(* IEC 61131-3 sources: plcassist-cli/packages/volt-lsp-iec/test-corpus/bakon-nano/Device/Plc Logic/Application/Library Manager/CAA Storage Imp, 116 files *)

(* ---- _3SSTORAGEVERSIONCONSTANTS.gvl ---- *)
VAR_GLOBAL
	_3SSTORAGE_VERSION_LARGEROREQUAL_3_5_5_0_ : INT := 0;
	_3SSTORAGE_VERSION_LARGEROREQUAL_3_5_11_10_ : INT := 0;
END_VAR

(* ---- GLOBALVARIABLES.gvl ---- *)
VAR_GLOBAL
	FACTORY : StorageFactory;
END_VAR

(* ---- _COLUMNGETBLOB.fun ---- *)
FUNCTION _COLUMNGETBLOB : STO.ERROR
VAR_INPUT
	HROW : ROW;
	IDCOLUMN : CAA.IDENT;
END_VAR
VAR_OUTPUT
	XNULL : BOOL;
END_VAR
VAR_IN_OUT
	BLOBVALUE : STO.STO_BLOB;
END_VAR
END_FUNCTION

(* ---- _COLUMNGETINT16.fun ---- *)
FUNCTION _COLUMNGETINT16 : STO.ERROR
VAR_INPUT
	HROW : ROW;
	IDCOLUMN : CAA.IDENT;
END_VAR
VAR_OUTPUT
	IVALUE : INT;
	XNULL : BOOL;
END_VAR
END_FUNCTION

(* ---- _COLUMNGETINT32.fun ---- *)
FUNCTION _COLUMNGETINT32 : STO.ERROR
VAR_INPUT
	HROW : ROW;
	IDCOLUMN : CAA.IDENT;
END_VAR
VAR_OUTPUT
	DIVALUE : DINT;
	XNULL : BOOL;
END_VAR
END_FUNCTION

(* ---- _COLUMNGETINT64.fun ---- *)
FUNCTION _COLUMNGETINT64 : STO.ERROR
VAR_INPUT
	HROW : ROW;
	IDCOLUMN : CAA.IDENT;
END_VAR
VAR_OUTPUT
	LIVALUE : LINT;
	XNULL : BOOL;
END_VAR
END_FUNCTION

(* ---- _COLUMNGETINT8.fun ---- *)
FUNCTION _COLUMNGETINT8 : STO.ERROR
VAR_INPUT
	HROW : ROW;
	IDCOLUMN : CAA.IDENT;
END_VAR
VAR_OUTPUT
	SIVALUE : SINT;
	XNULL : BOOL;
END_VAR
END_FUNCTION

(* ---- _COLUMNGETREAL4.fun ---- *)
FUNCTION _COLUMNGETREAL4 : STO.ERROR
VAR_INPUT
	HROW : ROW;
	IDCOLUMN : CAA.IDENT;
END_VAR
VAR_OUTPUT
	RVALUE : REAL;
	XNULL : BOOL;
END_VAR
END_FUNCTION

(* ---- _COLUMNGETREAL8.fun ---- *)
FUNCTION _COLUMNGETREAL8 : STO.ERROR
VAR_INPUT
	HROW : ROW;
	IDCOLUMN : CAA.IDENT;
END_VAR
VAR_OUTPUT
	LRVALUE : LREAL;
	XNULL : BOOL;
END_VAR
END_FUNCTION

(* ---- _COLUMNGETTEXT.fun ---- *)
FUNCTION _COLUMNGETTEXT : STO.ERROR
VAR_INPUT
	HROW : ROW;
	IDCOLUMN : CAA.IDENT;
END_VAR
VAR_OUTPUT
	XNULL : BOOL;
END_VAR
VAR_IN_OUT
	TXTVALUE : STO.STO_TEXT;
END_VAR
END_FUNCTION

(* ---- _COLUMNGETTYPE.fun ---- *)
FUNCTION _COLUMNGETTYPE : STO.COLUMN_TYPE
VAR_INPUT
	HROW : ROW;
	IDCOLUMN : CAA.IDENT;
END_VAR
VAR_OUTPUT
	EERROR : STO.ERROR;
END_VAR
END_FUNCTION

(* ---- _COLUMNSETBLOB.fun ---- *)
FUNCTION _COLUMNSETBLOB : STO.ERROR
VAR_INPUT
	HROW : ROW;
	IDCOLUMN : CAA.IDENT;
END_VAR
VAR_IN_OUT
	BLOBVALUE : STO.STO_BLOB;
END_VAR
END_FUNCTION

(* ---- _COLUMNSETINT16.fun ---- *)
FUNCTION _COLUMNSETINT16 : STO.ERROR
VAR_INPUT
	HROW : ROW;
	IDCOLUMN : CAA.IDENT;
	IVALUE : INT;
END_VAR
END_FUNCTION

(* ---- _COLUMNSETINT32.fun ---- *)
FUNCTION _COLUMNSETINT32 : STO.ERROR
VAR_INPUT
	HROW : ROW;
	IDCOLUMN : CAA.IDENT;
	DIVALUE : DINT;
END_VAR
END_FUNCTION

(* ---- _COLUMNSETINT64.fun ---- *)
FUNCTION _COLUMNSETINT64 : STO.ERROR
VAR_INPUT
	HROW : ROW;
	IDCOLUMN : CAA.IDENT;
	LIVALUE : LINT;
END_VAR
END_FUNCTION

(* ---- _COLUMNSETINT8.fun ---- *)
FUNCTION _COLUMNSETINT8 : STO.ERROR
VAR_INPUT
	HROW : ROW;
	IDCOLUMN : CAA.IDENT;
	SIVALUE : SINT;
END_VAR
END_FUNCTION

(* ---- _COLUMNSETNULL.fun ---- *)
FUNCTION _COLUMNSETNULL : STO.ERROR
VAR_INPUT
	HROW : ROW;
	IDCOLUMN : CAA.IDENT;
END_VAR
END_FUNCTION

(* ---- _COLUMNSETREAL4.fun ---- *)
FUNCTION _COLUMNSETREAL4 : STO.ERROR
VAR_INPUT
	HROW : ROW;
	IDCOLUMN : CAA.IDENT;
	RVALUE : REAL;
END_VAR
END_FUNCTION

(* ---- _COLUMNSETREAL8.fun ---- *)
FUNCTION _COLUMNSETREAL8 : STO.ERROR
VAR_INPUT
	HROW : ROW;
	IDCOLUMN : CAA.IDENT;
	LRVALUE : LREAL;
END_VAR
END_FUNCTION

(* ---- _COLUMNSETTEXT.fun ---- *)
FUNCTION _COLUMNSETTEXT : STO.ERROR
VAR_INPUT
	HROW : ROW;
	IDCOLUMN : CAA.IDENT;
END_VAR
VAR_IN_OUT
	TXTVALUE : STO.STO_TEXT;
END_VAR
END_FUNCTION

(* ---- _COLUMNUPDATEBLOB.fun ---- *)
FUNCTION _COLUMNUPDATEBLOB : STO.ERROR
VAR_INPUT
	HROW : ROW;
	IDCOLUMN : CAA.IDENT;
END_VAR
VAR_IN_OUT
	BLOBVALUE : STO.STO_BLOB;
	XNULL : BOOL;
END_VAR
END_FUNCTION

(* ---- _COLUMNUPDATEINT16.fun ---- *)
FUNCTION _COLUMNUPDATEINT16 : STO.ERROR
VAR_INPUT
	HROW : ROW;
	IDCOLUMN : CAA.IDENT;
END_VAR
VAR_IN_OUT
	IVALUE : INT;
	XNULL : BOOL;
END_VAR
END_FUNCTION

(* ---- _COLUMNUPDATEINT32.fun ---- *)
FUNCTION _COLUMNUPDATEINT32 : STO.ERROR
VAR_INPUT
	HROW : ROW;
	IDCOLUMN : CAA.IDENT;
END_VAR
VAR_IN_OUT
	DIVALUE : DINT;
	XNULL : BOOL;
END_VAR
END_FUNCTION

(* ---- _COLUMNUPDATEINT64.fun ---- *)
FUNCTION _COLUMNUPDATEINT64 : STO.ERROR
VAR_INPUT
	HROW : ROW;
	IDCOLUMN : CAA.IDENT;
END_VAR
VAR_IN_OUT
	LIVALUE : LINT;
	XNULL : BOOL;
END_VAR
END_FUNCTION

(* ---- _COLUMNUPDATEINT8.fun ---- *)
FUNCTION _COLUMNUPDATEINT8 : STO.ERROR
VAR_INPUT
	HROW : ROW;
	IDCOLUMN : CAA.IDENT;
END_VAR
VAR_IN_OUT
	SIVALUE : SINT;
	XNULL : BOOL;
END_VAR
END_FUNCTION

(* ---- _COLUMNUPDATEREAL4.fun ---- *)
FUNCTION _COLUMNUPDATEREAL4 : STO.ERROR
VAR_INPUT
	HROW : ROW;
	IDCOLUMN : CAA.IDENT;
END_VAR
VAR_IN_OUT
	RVALUE : REAL;
	XNULL : BOOL;
END_VAR
END_FUNCTION

(* ---- _COLUMNUPDATEREAL8.fun ---- *)
FUNCTION _COLUMNUPDATEREAL8 : STO.ERROR
VAR_INPUT
	HROW : ROW;
	IDCOLUMN : CAA.IDENT;
END_VAR
VAR_IN_OUT
	LRVALUE : LREAL;
	XNULL : BOOL;
END_VAR
END_FUNCTION

(* ---- _COLUMNUPDATETEXT.fun ---- *)
FUNCTION _COLUMNUPDATETEXT : STO.ERROR
VAR_INPUT
	HROW : ROW;
	IDCOLUMN : CAA.IDENT;
END_VAR
VAR_IN_OUT
	TXTVALUE : STO.STO_TEXT;
	XNULL : BOOL;
END_VAR
END_FUNCTION

(* ---- _CURSORCLOSE.fun ---- *)
FUNCTION _CURSORCLOSE : STO.ERROR
VAR_INPUT
	HCURSOR : CURSOR;
END_VAR
END_FUNCTION

(* ---- _CURSORGETCURRENTROW.fun ---- *)
FUNCTION _CURSORGETCURRENTROW : ROW
VAR_INPUT
	HCURSOR : CURSOR;
END_VAR
VAR_OUTPUT
	EERROR : STO.ERROR;
END_VAR
END_FUNCTION

(* ---- _CURSORGETINDEXID.fun ---- *)
FUNCTION _CURSORGETINDEXID : CAA.IDENT
VAR_INPUT
	HCURSOR : CURSOR;
END_VAR
VAR_OUTPUT
	EERROR : STO.ERROR;
END_VAR
END_FUNCTION

(* ---- _CURSORGETSTORAGE.fun ---- *)
FUNCTION _CURSORGETSTORAGE : STORAGE_TYPE
VAR_INPUT
	HCURSOR : CURSOR;
END_VAR
VAR_OUTPUT
	EERROR : STO.ERROR;
END_VAR
END_FUNCTION

(* ---- _CURSORGETTABLE.fun ---- *)
FUNCTION _CURSORGETTABLE : TABLE
VAR_INPUT
	HCURSOR : CURSOR;
END_VAR
VAR_OUTPUT
	EERROR : STO.ERROR;
END_VAR
END_FUNCTION

(* ---- _CURSORISREADONLY.fun ---- *)
FUNCTION _CURSORISREADONLY : BOOL
VAR_INPUT
	HCURSOR : CURSOR;
END_VAR
VAR_OUTPUT
	EERROR : STO.ERROR;
END_VAR
END_FUNCTION

(* ---- _CURSORMOVE.fun ---- *)
FUNCTION _CURSORMOVE : STO.ERROR
VAR_INPUT
	HCURSOR : CURSOR;
	EDIRECTION : STO.DIRECTION;
END_VAR
END_FUNCTION

(* ---- _CURSOROPEN.fun ---- *)
FUNCTION _CURSOROPEN : CURSOR
VAR_INPUT
	HTABLE : TABLE;
	IDINDEX : CAA.IDENT;
	XREADONLY : BOOL;
END_VAR
VAR_OUTPUT
	EERROR : STO.ERROR;
END_VAR
END_FUNCTION

(* ---- _CURSORSEARCHINT16.fun ---- *)
FUNCTION _CURSORSEARCHINT16 : STO.ERROR
VAR_INPUT
	HCURSOR : CURSOR;
	IVALUE : INT;
END_VAR
END_FUNCTION

(* ---- _CURSORSEARCHINT32.fun ---- *)
FUNCTION _CURSORSEARCHINT32 : STO.ERROR
VAR_INPUT
	HCURSOR : CURSOR;
	DIVALUE : DINT;
END_VAR
END_FUNCTION

(* ---- _CURSORSEARCHINT64.fun ---- *)
FUNCTION _CURSORSEARCHINT64 : STO.ERROR
VAR_INPUT
	HCURSOR : CURSOR;
	LIVALUE : LINT;
END_VAR
END_FUNCTION

(* ---- _CURSORSEARCHINT8.fun ---- *)
FUNCTION _CURSORSEARCHINT8 : STO.ERROR
VAR_INPUT
	HCURSOR : CURSOR;
	SIVALUE : SINT;
END_VAR
END_FUNCTION

(* ---- _CURSORSEARCHNULL.fun ---- *)
FUNCTION _CURSORSEARCHNULL : STO.ERROR
VAR_INPUT
	HCURSOR : CURSOR;
END_VAR
END_FUNCTION

(* ---- _CURSORSEARCHREAL4.fun ---- *)
FUNCTION _CURSORSEARCHREAL4 : STO.ERROR
VAR_INPUT
	HCURSOR : CURSOR;
	RVALUE : REAL;
END_VAR
END_FUNCTION

(* ---- _CURSORSEARCHREAL8.fun ---- *)
FUNCTION _CURSORSEARCHREAL8 : STO.ERROR
VAR_INPUT
	HCURSOR : CURSOR;
	LRVALUE : LREAL;
END_VAR
END_FUNCTION

(* ---- _CURSORSEARCHROWID.fun ---- *)
FUNCTION _CURSORSEARCHROWID : STO.ERROR
VAR_INPUT
	HCURSOR : CURSOR;
	IDROW : CAA.IDENT;
END_VAR
END_FUNCTION

(* ---- _CURSORSEARCHROWID2.fun ---- *)
FUNCTION _CURSORSEARCHROWID2 : STO.ERROR
VAR_INPUT
	HCURSOR : CURSOR;
	IDROW : LINT;
END_VAR
END_FUNCTION

(* ---- _CURSORSEARCHTEXT.fun ---- *)
FUNCTION _CURSORSEARCHTEXT : STO.ERROR
VAR_INPUT
	HCURSOR : CURSOR;
END_VAR
VAR_IN_OUT
	TXTVALUE : STO.STO_TEXT;
END_VAR
END_FUNCTION

(* ---- _ROWCLEAR.fun ---- *)
FUNCTION _ROWCLEAR : STO.ERROR
VAR_INPUT
	HROW : ROW;
END_VAR
END_FUNCTION

(* ---- _ROWCREATE.fun ---- *)
FUNCTION _ROWCREATE : ROW
VAR_INPUT
	HTABLE : TABLE;
END_VAR
VAR_OUTPUT
	EERROR : STO.ERROR;
END_VAR
END_FUNCTION

(* ---- _ROWDELETE.fun ---- *)
FUNCTION _ROWDELETE : STO.ERROR
VAR_INPUT
	HTABLE : TABLE;
	IDROW : CAA.IDENT;
END_VAR
END_FUNCTION

(* ---- _ROWDELETE2.fun ---- *)
FUNCTION _ROWDELETE2 : STO.ERROR
VAR_INPUT
	HTABLE : TABLE;
	IDROW : LINT;
END_VAR
END_FUNCTION

(* ---- _ROWDUPLICATE.fun ---- *)
FUNCTION _ROWDUPLICATE : ROW
VAR_INPUT
	HTABLE : TABLE;
	IDROW : CAA.IDENT;
END_VAR
VAR_OUTPUT
	EERROR : STO.ERROR;
END_VAR
END_FUNCTION

(* ---- _ROWGETHASCHANGED.fun ---- *)
FUNCTION _ROWGETHASCHANGED : BOOL
VAR_INPUT
	HROW : ROW;
END_VAR
VAR_OUTPUT
	EERROR : STO.ERROR;
END_VAR
END_FUNCTION

(* ---- _ROWGETID.fun ---- *)
FUNCTION _ROWGETID : CAA.IDENT
VAR_INPUT
	HROW : ROW;
END_VAR
VAR_OUTPUT
	EERROR : STO.ERROR;
END_VAR
END_FUNCTION

(* ---- _ROWGETID2.fun ---- *)
FUNCTION _ROWGETID2 : LINT
VAR_INPUT
	HROW : ROW;
END_VAR
VAR_OUTPUT
	EERROR : STO.ERROR;
END_VAR
END_FUNCTION

(* ---- _ROWGETNUMOFCOLUMNS.fun ---- *)
FUNCTION _ROWGETNUMOFCOLUMNS : CAA.COUNT
VAR_INPUT
	HROW : ROW;
END_VAR
VAR_OUTPUT
	EERROR : STO.ERROR;
END_VAR
END_FUNCTION

(* ---- _ROWGETSTORAGE.fun ---- *)
FUNCTION _ROWGETSTORAGE : STORAGE_TYPE
VAR_INPUT
	HROW : ROW;
END_VAR
VAR_OUTPUT
	EERROR : STO.ERROR;
END_VAR
END_FUNCTION

(* ---- _ROWGETTABLE.fun ---- *)
FUNCTION _ROWGETTABLE : TABLE
VAR_INPUT
	HROW : ROW;
END_VAR
VAR_OUTPUT
	EERROR : STO.ERROR;
END_VAR
END_FUNCTION

(* ---- _ROWINSERT.fun ---- *)
FUNCTION _ROWINSERT : CAA.IDENT
VAR_INPUT
	HROW : ROW;
END_VAR
VAR_OUTPUT
	EERROR : STO.ERROR;
END_VAR
END_FUNCTION

(* ---- _ROWRELEASE.fun ---- *)
FUNCTION _ROWRELEASE : STO.ERROR
VAR_INPUT
	HROW : ROW;
END_VAR
END_FUNCTION

(* ---- _ROWSELECT.fun ---- *)
FUNCTION _ROWSELECT : ROW
VAR_INPUT
	HTABLE : TABLE;
	IDROW : CAA.IDENT;
END_VAR
VAR_OUTPUT
	EERROR : STO.ERROR;
END_VAR
END_FUNCTION

(* ---- _ROWUPDATE.fun ---- *)
FUNCTION _ROWUPDATE : STO.ERROR
VAR_INPUT
	HROW : ROW;
END_VAR
END_FUNCTION

(* ---- _SAVEPOINTGETSTORAGE.fun ---- *)
FUNCTION _SAVEPOINTGETSTORAGE : STORAGE_TYPE
VAR_INPUT
	HSAVEPOINT : SAVEPOINT;
END_VAR
VAR_OUTPUT
	EERROR : STO.ERROR;
END_VAR
END_FUNCTION

(* ---- _SAVEPOINTGETTRANSACTION.fun ---- *)
FUNCTION _SAVEPOINTGETTRANSACTION : TRANSACTION
VAR_INPUT
	HSAVEPOINT : SAVEPOINT;
END_VAR
VAR_OUTPUT
	EERROR : STO.ERROR;
END_VAR
END_FUNCTION

(* ---- _SAVEPOINTRELEASE.fun ---- *)
FUNCTION _SAVEPOINTRELEASE : STO.ERROR
VAR_INPUT
	HSAVEPOINT : SAVEPOINT;
END_VAR
END_FUNCTION

(* ---- _SAVEPOINTROLLBACK.fun ---- *)
FUNCTION _SAVEPOINTROLLBACK : STO.ERROR
VAR_INPUT
	HSAVEPOINT : SAVEPOINT;
END_VAR
END_FUNCTION

(* ---- _STORAGECLEAR.fun ---- *)
FUNCTION _STORAGECLEAR : STO.ERROR
VAR_INPUT
	HSTORAGE : STORAGE_TYPE;
END_VAR
END_FUNCTION

(* ---- _STORAGECLOSE.fun ---- *)
FUNCTION _STORAGECLOSE : STO.ERROR
VAR_INPUT
	HSTORAGE : STORAGE_TYPE;
END_VAR
END_FUNCTION

(* ---- _STORAGEEXECUTESTATEMENT.fun ---- *)
FUNCTION _STORAGEEXECUTESTATEMENT : STO.ERROR
VAR_INPUT
	HSTORAGE : STORAGE_TYPE;
END_VAR
VAR_IN_OUT
	SSTATEMENT : STO.SQLSTATEMENT;
END_VAR
END_FUNCTION

(* ---- _STORAGEGETENCODING.fun ---- *)
FUNCTION _STORAGEGETENCODING : STO.ENCODING
VAR_INPUT
	HSTORAGE : STORAGE_TYPE;
END_VAR
VAR_OUTPUT
	EERROR : STO.ERROR;
END_VAR
END_FUNCTION

(* ---- _STORAGEGETINDEXID.fun ---- *)
FUNCTION _STORAGEGETINDEXID : STO.ERROR
VAR_INPUT
	HSTORAGE : STORAGE_TYPE;
END_VAR
VAR_OUTPUT
	IDINDEX : CAA.IDENT;
END_VAR
VAR_IN_OUT
	SINDEX : STRING;
	STABLE : STRING;
END_VAR
END_FUNCTION

(* ---- _STORAGEGETLOCKINGSTATE.fun ---- *)
FUNCTION _STORAGEGETLOCKINGSTATE : STO.LOCKING_STATE
VAR_INPUT
	HSTORAGE : STORAGE_TYPE;
END_VAR
VAR_OUTPUT
	EERROR : STO.ERROR;
END_VAR
END_FUNCTION

(* ---- _STORAGEGETMETRICS.fun ---- *)
FUNCTION _STORAGEGETMETRICS : STO.ERROR
VAR_INPUT
	HSTORAGE : STORAGE_TYPE;
END_VAR
VAR_IN_OUT
	MMETRICS : STO.STO_METRICS;
END_VAR
END_FUNCTION

(* ---- _STORAGEGETNUMOFTABLES.fun ---- *)
FUNCTION _STORAGEGETNUMOFTABLES : CAA.COUNT
VAR_INPUT
	HSTORAGE : STORAGE_TYPE;
END_VAR
VAR_OUTPUT
	EERROR : STO.ERROR;
END_VAR
END_FUNCTION

(* ---- _STORAGEGETPATH.fun ---- *)
FUNCTION _STORAGEGETPATH : STO.ERROR
VAR_INPUT
	HSTORAGE : STORAGE_TYPE;
END_VAR
VAR_IN_OUT
	SPATH : CAA.FILENAME;
END_VAR
END_FUNCTION

(* ---- _STORAGEGETSCHEMAVERSION.fun ---- *)
FUNCTION _STORAGEGETSCHEMAVERSION : DINT
VAR_INPUT
	HSTORAGE : STORAGE_TYPE;
END_VAR
VAR_OUTPUT
	EERROR : STO.ERROR;
END_VAR
END_FUNCTION

(* ---- _STORAGEGETSTORAGEVERSION.fun ---- *)
FUNCTION _STORAGEGETSTORAGEVERSION : DINT
VAR_INPUT
	HSTORAGE : STORAGE_TYPE;
END_VAR
VAR_OUTPUT
	EERROR : STO.ERROR;
END_VAR
END_FUNCTION

(* ---- _STORAGEGETTABLEID.fun ---- *)
FUNCTION _STORAGEGETTABLEID : STO.ERROR
VAR_INPUT
	HSTORAGE : STORAGE_TYPE;
END_VAR
VAR_OUTPUT
	IDTABLE : CAA.IDENT;
END_VAR
VAR_IN_OUT
	STABLE : STRING;
END_VAR
END_FUNCTION

(* ---- _STORAGEGETUSERVERSION.fun ---- *)
FUNCTION _STORAGEGETUSERVERSION : DINT
VAR_INPUT
	HSTORAGE : STORAGE_TYPE;
END_VAR
VAR_OUTPUT
	EERROR : STO.ERROR;
END_VAR
END_FUNCTION

(* ---- _STORAGEISREADONLY.fun ---- *)
FUNCTION _STORAGEISREADONLY : BOOL
VAR_INPUT
	HSTORAGE : STORAGE_TYPE;
END_VAR
VAR_OUTPUT
	EERROR : STO.ERROR;
END_VAR
END_FUNCTION

(* ---- _STORAGEOPENFILE.fun ---- *)
FUNCTION _STORAGEOPENFILE : STORAGE_TYPE
VAR_INPUT
	SPATH : CAA.FILENAME;
	XREADONLY : BOOL := FALSE;
END_VAR
VAR_OUTPUT
	EERROR : STO.ERROR;
END_VAR
END_FUNCTION

(* ---- _STORAGEREORG.fun ---- *)
FUNCTION _STORAGEREORG : STO.ERROR
VAR_INPUT
	HSTORAGE : STORAGE_TYPE;
END_VAR
END_FUNCTION

(* ---- _TABLECLEAR.fun ---- *)
FUNCTION _TABLECLEAR : STO.ERROR
VAR_INPUT
	HTABLE : TABLE;
END_VAR
END_FUNCTION

(* ---- _TABLECLOSE.fun ---- *)
FUNCTION _TABLECLOSE : STO.ERROR
VAR_INPUT
	HTABLE : TABLE;
END_VAR
END_FUNCTION

(* ---- _TABLEGETID.fun ---- *)
FUNCTION _TABLEGETID : CAA.IDENT
VAR_INPUT
	HTABLE : TABLE;
END_VAR
VAR_OUTPUT
	EERROR : STO.ERROR;
END_VAR
END_FUNCTION

(* ---- _TABLEGETMINMAXROWIDS.fun ---- *)
FUNCTION _TABLEGETMINMAXROWIDS : STO.ERROR
VAR_INPUT
	HTABLE : TABLE;
END_VAR
VAR_OUTPUT
	IDROWMIN : LINT;
	IDROWMAX : LINT;
END_VAR
END_FUNCTION

(* ---- _TABLEGETNUMOFCOLUMNS.fun ---- *)
FUNCTION _TABLEGETNUMOFCOLUMNS : CAA.COUNT
VAR_INPUT
	HTABLE : TABLE;
END_VAR
VAR_OUTPUT
	EERROR : STO.ERROR;
END_VAR
END_FUNCTION

(* ---- _TABLEGETNUMOFINDEXES.fun ---- *)
FUNCTION _TABLEGETNUMOFINDEXES : CAA.COUNT
VAR_INPUT
	HTABLE : TABLE;
END_VAR
VAR_OUTPUT
	EERROR : STO.ERROR;
END_VAR
END_FUNCTION

(* ---- _TABLEGETNUMOFROWS.fun ---- *)
FUNCTION _TABLEGETNUMOFROWS : CAA.COUNT
VAR_INPUT
	HTABLE : TABLE;
END_VAR
VAR_OUTPUT
	EERROR : STO.ERROR;
END_VAR
END_FUNCTION

(* ---- _TABLEGETSTORAGE.fun ---- *)
FUNCTION _TABLEGETSTORAGE : STORAGE_TYPE
VAR_INPUT
	HTABLE : TABLE;
END_VAR
VAR_OUTPUT
	EERROR : STO.ERROR;
END_VAR
END_FUNCTION

(* ---- _TABLEOPEN.fun ---- *)
FUNCTION _TABLEOPEN : TABLE
VAR_INPUT
	HSTORAGE : STORAGE_TYPE;
	IDTABLE : CAA.IDENT;
END_VAR
VAR_OUTPUT
	EERROR : STO.ERROR;
END_VAR
END_FUNCTION

(* ---- _TRANSACTIONBEGIN.fun ---- *)
FUNCTION _TRANSACTIONBEGIN : TRANSACTION
VAR_INPUT
	HSTORAGE : STORAGE_TYPE;
	EMODE : STO.TRANSACTION_MODE;
END_VAR
VAR_OUTPUT
	EERROR : STO.ERROR;
END_VAR
END_FUNCTION

(* ---- _TRANSACTIONCOMMIT.fun ---- *)
FUNCTION _TRANSACTIONCOMMIT : STO.ERROR
VAR_INPUT
	HTRANSACTION : TRANSACTION;
END_VAR
END_FUNCTION

(* ---- _TRANSACTIONGETSTORAGE.fun ---- *)
FUNCTION _TRANSACTIONGETSTORAGE : STORAGE_TYPE
VAR_INPUT
	HTRANSACTION : TRANSACTION;
END_VAR
VAR_OUTPUT
	EERROR : STO.ERROR;
END_VAR
END_FUNCTION

(* ---- _TRANSACTIONROLLBACK.fun ---- *)
FUNCTION _TRANSACTIONROLLBACK : STO.ERROR
VAR_INPUT
	HTRANSACTION : TRANSACTION;
END_VAR
END_FUNCTION

(* ---- _TRANSACTIONSETSAVEPOINT.fun ---- *)
FUNCTION _TRANSACTIONSETSAVEPOINT : SAVEPOINT
VAR_INPUT
	HTRANSACTION : TRANSACTION;
END_VAR
VAR_OUTPUT
	EERROR : STO.ERROR;
END_VAR
END_FUNCTION

(* ---- _UTILITYGETCURRENTDATEANDTIME.fun ---- *)
FUNCTION _UTILITYGETCURRENTDATEANDTIME : STO.INT64
VAR_INPUT
	HSTORAGE : STORAGE_TYPE;
END_VAR
VAR_OUTPUT
	EERROR : STO.ERROR;
END_VAR
END_FUNCTION

(* ---- _UTILITYRANDOMNESS.fun ---- *)
FUNCTION _UTILITYRANDOMNESS : STO.ERROR
VAR_INPUT
	HSTORAGE : STORAGE_TYPE;
	SZSIZE : CAA.SIZE;
	PDATA : CAA.PVOID;
END_VAR
END_FUNCTION

(* ---- CURSORIMP.fb ---- *)
FUNCTION_BLOCK CURSORIMP EXTENDS InstanceBase
VAR
	_HHANDLE : CAA.HANDLE;
	_ITFTABLE : STO.ITable;
	_EERROR : STO.ERROR;
	CURSORCURRENTROW : STO.IRow;
	CURSORINDEXID : CAA.IDENT;
	CURSORISREADONLY : BOOL;
	CURSORSTORAGE : STO.IStorage;
	CURSORTABLE : STO.ITable;
	LASTERROR : STO.ERROR;
END_VAR
END_FUNCTION_BLOCK

METHOD CURSORCLOSE : STO.ERROR
END_METHOD

METHOD CURSORMOVE : STO.ERROR
VAR_INPUT
	EDIRECTION : STO.DIRECTION;
END_VAR
END_METHOD

METHOD CURSORSEARCHROWID : STO.ERROR
VAR_INPUT
	IDROW : CAA.IDENT;
END_VAR
END_METHOD

METHOD CURSORSEARCHROWID2 : STO.ERROR
VAR_INPUT
	IDROW : LINT;
END_VAR
END_METHOD

METHOD CURSORSEARCH_DINT : STO.ERROR
VAR_INPUT
	DIVALUE : DINT;
END_VAR
END_METHOD

METHOD CURSORSEARCH_INT : STO.ERROR
VAR_INPUT
	IVALUE : INT;
END_VAR
END_METHOD

METHOD CURSORSEARCH_LINT : STO.ERROR
VAR_INPUT
	LIVALUE : LINT;
END_VAR
END_METHOD

METHOD CURSORSEARCH_LREAL : STO.ERROR
VAR_INPUT
	LRVALUE : LREAL;
END_VAR
END_METHOD

METHOD CURSORSEARCH_NULL : STO.ERROR
END_METHOD

METHOD CURSORSEARCH_REAL : STO.ERROR
VAR_INPUT
	RVALUE : REAL;
END_VAR
END_METHOD

METHOD CURSORSEARCH_SINT : STO.ERROR
VAR_INPUT
	SIVALUE : SINT;
END_VAR
END_METHOD

METHOD CURSORSEARCH_TEXT : STO.ERROR
VAR_IN_OUT
	TXTVALUE : STO.TEXT;
END_VAR
END_METHOD

METHOD PRVINSTINIT : FBF.ERROR
VAR_INPUT
	ITFDATA : FBF.IData;
END_VAR
END_METHOD

(* ---- CURSORIMPFACTORY.fb ---- *)
FUNCTION_BLOCK CURSORIMPFACTORY EXTENDS FactoryBase
VAR
	PRVINSTCOUNT : CAA.COUNT;
	PRVINSTPOOLEXTENDSFACTOR : USINT;
	PRVINSTSIZE : CAA.SIZE;
END_VAR
END_FUNCTION_BLOCK

METHOD CREATE : POINTER TO CursorImp
VAR_INPUT
	ITFDATA : FBF.IData;
END_VAR
VAR_OUTPUT
	EERROR : FBF.ERROR;
END_VAR
END_METHOD

(* ---- INITDATA.fb ---- *)
FUNCTION_BLOCK INITDATA EXTENDS InstanceData
VAR_INPUT
	HHANDLE : CAA.HANDLE;
END_VAR
END_FUNCTION_BLOCK

(* ---- INITSTORAGEDATA.fb ---- *)
FUNCTION_BLOCK INITSTORAGEDATA EXTENDS InitData
VAR_INPUT
	ITFSTORAGE : STO.IStorage;
END_VAR
END_FUNCTION_BLOCK

(* ---- INITTABLEDATA.fb ---- *)
FUNCTION_BLOCK INITTABLEDATA EXTENDS InitData
VAR_INPUT
	ITFTABLE : STO.ITable;
END_VAR
END_FUNCTION_BLOCK

(* ---- INITTRANSACTIONDATA.fb ---- *)
FUNCTION_BLOCK INITTRANSACTIONDATA EXTENDS InitData
VAR_INPUT
	ITFTRANSACTION : STO.ITransaction;
END_VAR
END_FUNCTION_BLOCK

(* ---- ROWBASEIMP.fb ---- *)
FUNCTION_BLOCK ROWBASEIMP EXTENDS InstanceBase
VAR
	_HHANDLE : CAA.HANDLE;
	_ITFTABLE : STO.ITable;
	ROWNUMOFCOLUMNS : CAA.COUNT;
	ROWSTORAGE : STO.IStorage;
	ROWTABLE : STO.ITable;
END_VAR
END_FUNCTION_BLOCK

METHOD COLUMNGETTYPE : STO.COLUMN_TYPE
VAR_INPUT
	IDCOLUMN : CAA.IDENT;
END_VAR
VAR_OUTPUT
	EERROR : STO.ERROR;
END_VAR
END_METHOD

METHOD COLUMNGET_BLOB : STO.ERROR
VAR_INPUT
	IDCOLUMN : CAA.IDENT;
END_VAR
VAR_OUTPUT
	XNULL : BOOL;
END_VAR
VAR_IN_OUT
	BLOBVALUE : STO.BLOB;
END_VAR
END_METHOD

METHOD COLUMNGET_DINT : STO.ERROR
VAR_INPUT
	IDCOLUMN : CAA.IDENT;
END_VAR
VAR_OUTPUT
	DIVALUE : DINT;
	XNULL : BOOL;
END_VAR
END_METHOD

METHOD COLUMNGET_INT : STO.ERROR
VAR_INPUT
	IDCOLUMN : CAA.IDENT;
END_VAR
VAR_OUTPUT
	IVALUE : INT;
	XNULL : BOOL;
END_VAR
END_METHOD

METHOD COLUMNGET_LINT : STO.ERROR
VAR_INPUT
	IDCOLUMN : CAA.IDENT;
END_VAR
VAR_OUTPUT
	LIVALUE : LINT;
	XNULL : BOOL;
END_VAR
END_METHOD

METHOD COLUMNGET_LREAL : STO.ERROR
VAR_INPUT
	IDCOLUMN : CAA.IDENT;
END_VAR
VAR_OUTPUT
	LRVALUE : LREAL;
	XNULL : BOOL;
END_VAR
END_METHOD

METHOD COLUMNGET_REAL : STO.ERROR
VAR_INPUT
	IDCOLUMN : CAA.IDENT;
END_VAR
VAR_OUTPUT
	RVALUE : REAL;
	XNULL : BOOL;
END_VAR
END_METHOD

METHOD COLUMNGET_SINT : STO.ERROR
VAR_INPUT
	IDCOLUMN : CAA.IDENT;
END_VAR
VAR_OUTPUT
	SIVALUE : SINT;
	XNULL : BOOL;
END_VAR
END_METHOD

METHOD COLUMNGET_TEXT : STO.ERROR
VAR_INPUT
	IDCOLUMN : CAA.IDENT;
END_VAR
VAR_OUTPUT
	XNULL : BOOL;
END_VAR
VAR_IN_OUT
	TXTVALUE : STO.TEXT;
END_VAR
END_METHOD

METHOD COLUMNSET_BLOB : STO.ERROR
VAR_INPUT
	IDCOLUMN : CAA.IDENT;
END_VAR
VAR_IN_OUT
	BLOBVALUE : STO.BLOB;
END_VAR
END_METHOD

METHOD COLUMNSET_DINT : STO.ERROR
VAR_INPUT
	IDCOLUMN : CAA.IDENT;
	DIVALUE : DINT;
END_VAR
END_METHOD

METHOD COLUMNSET_INT : STO.ERROR
VAR_INPUT
	IDCOLUMN : CAA.IDENT;
	IVALUE : INT;
END_VAR
END_METHOD

METHOD COLUMNSET_LINT : STO.ERROR
VAR_INPUT
	IDCOLUMN : CAA.IDENT;
	LIVALUE : LINT;
END_VAR
END_METHOD

METHOD COLUMNSET_LREAL : STO.ERROR
VAR_INPUT
	IDCOLUMN : CAA.IDENT;
	LRVALUE : LREAL;
END_VAR
END_METHOD

METHOD COLUMNSET_NULL : STO.ERROR
VAR_INPUT
	IDCOLUMN : CAA.IDENT;
END_VAR
END_METHOD

METHOD COLUMNSET_REAL : STO.ERROR
VAR_INPUT
	IDCOLUMN : CAA.IDENT;
	RVALUE : REAL;
END_VAR
END_METHOD

METHOD COLUMNSET_SINT : STO.ERROR
VAR_INPUT
	IDCOLUMN : CAA.IDENT;
	SIVALUE : SINT;
END_VAR
END_METHOD

METHOD COLUMNSET_TEXT : STO.ERROR
VAR_INPUT
	IDCOLUMN : CAA.IDENT;
END_VAR
VAR_IN_OUT
	TXTVALUE : STO.TEXT;
END_VAR
END_METHOD

METHOD COLUMNUPDATE_BLOB : STO.ERROR
VAR_INPUT
	IDCOLUMN : CAA.IDENT;
END_VAR
VAR_IN_OUT
	BLOBVALUE : STO.BLOB;
	XNULL : BOOL;
END_VAR
END_METHOD

METHOD COLUMNUPDATE_DINT : STO.ERROR
VAR_INPUT
	IDCOLUMN : CAA.IDENT;
END_VAR
VAR_IN_OUT
	DIVALUE : DINT;
	XNULL : BOOL;
END_VAR
END_METHOD

METHOD COLUMNUPDATE_INT : STO.ERROR
VAR_INPUT
	IDCOLUMN : CAA.IDENT;
END_VAR
VAR_IN_OUT
	IVALUE : INT;
	XNULL : BOOL;
END_VAR
END_METHOD

METHOD COLUMNUPDATE_LINT : STO.ERROR
VAR_INPUT
	IDCOLUMN : CAA.IDENT;
END_VAR
VAR_IN_OUT
	LIVALUE : LINT;
	XNULL : BOOL;
END_VAR
END_METHOD

METHOD COLUMNUPDATE_LREAL : STO.ERROR
VAR_INPUT
	IDCOLUMN : CAA.IDENT;
END_VAR
VAR_IN_OUT
	LRVALUE : LREAL;
	XNULL : BOOL;
END_VAR
END_METHOD

METHOD COLUMNUPDATE_REAL : STO.ERROR
VAR_INPUT
	IDCOLUMN : CAA.IDENT;
END_VAR
VAR_IN_OUT
	RVALUE : REAL;
	XNULL : BOOL;
END_VAR
END_METHOD

METHOD COLUMNUPDATE_SINT : STO.ERROR
VAR_INPUT
	IDCOLUMN : CAA.IDENT;
END_VAR
VAR_IN_OUT
	SIVALUE : SINT;
	XNULL : BOOL;
END_VAR
END_METHOD

METHOD COLUMNUPDATE_TEXT : STO.ERROR
VAR_INPUT
	IDCOLUMN : CAA.IDENT;
END_VAR
VAR_IN_OUT
	TXTVALUE : STO.TEXT;
	XNULL : BOOL;
END_VAR
END_METHOD

METHOD ROWCLEAR : STO.ERROR
END_METHOD

METHOD ROWRELEASE : STO.ERROR
END_METHOD

METHOD PRVINSTINIT : FBF.ERROR
VAR_INPUT
	ITFDATA : FBF.IData;
END_VAR
END_METHOD

(* ---- ROWIMP.fb ---- *)
FUNCTION_BLOCK ROWIMP EXTENDS RowBaseImp
VAR
	EERROR : INT;
	_EERROR : STO.ERROR;
	LASTERROR : STO.ERROR;
	ROWHASCHANGED : BOOL;
	ROWID : CAA.IDENT;
END_VAR
END_FUNCTION_BLOCK

METHOD GETROWID : STO.ERROR
VAR_OUTPUT
	IDROW : LINT;
END_VAR
END_METHOD

METHOD ROWUPDATE : STO.ERROR
END_METHOD

(* ---- ROWIMPFACTORY.fb ---- *)
FUNCTION_BLOCK ROWIMPFACTORY EXTENDS FactoryBase
VAR
	PRVINSTCOUNT : CAA.COUNT;
	PRVINSTPOOLEXTENDSFACTOR : USINT;
	PRVINSTSIZE : CAA.SIZE;
END_VAR
END_FUNCTION_BLOCK

METHOD CREATE : POINTER TO RowImp
VAR_INPUT
	ITFDATA : FBF.IData;
END_VAR
VAR_OUTPUT
	EERROR : FBF.ERROR;
END_VAR
END_METHOD

(* ---- ROWPLANCHETIMP.fb ---- *)
FUNCTION_BLOCK ROWPLANCHETIMP EXTENDS RowBaseImp
END_FUNCTION_BLOCK

METHOD ROWINSERT : CAA.IDENT
VAR_OUTPUT
	EERROR : STO.ERROR;
END_VAR
END_METHOD

(* ---- ROWPLANCHETIMPFACTORY.fb ---- *)
FUNCTION_BLOCK ROWPLANCHETIMPFACTORY EXTENDS FactoryBase
VAR
	PRVINSTCOUNT : CAA.COUNT;
	PRVINSTPOOLEXTENDSFACTOR : USINT;
	PRVINSTSIZE : CAA.SIZE;
END_VAR
END_FUNCTION_BLOCK

METHOD CREATE : POINTER TO RowPlanchetImp
VAR_INPUT
	ITFDATA : FBF.IData;
END_VAR
VAR_OUTPUT
	EERROR : FBF.ERROR;
END_VAR
END_METHOD

(* ---- SAVEPOINTIMP.fb ---- *)
FUNCTION_BLOCK SAVEPOINTIMP EXTENDS InstanceBase
VAR
	_HHANDLE : CAA.HANDLE;
	_ITFTRANSACTION : STO.ITransaction;
	SAVEPOINTSTORAGE : STO.ISTorage;
	SAVEPOINTTRANSACTION : STO.ITransaction;
END_VAR
END_FUNCTION_BLOCK

METHOD SAVEPOINTROLLBACK : STO.ERROR
END_METHOD

METHOD SAVEPOINTRELEASE : STO.ERROR
END_METHOD

METHOD PRVINSTINIT : FBF.ERROR
VAR_INPUT
	ITFDATA : FBF.IData;
END_VAR
END_METHOD

(* ---- SAVEPOINTIMPFACTORY.fb ---- *)
FUNCTION_BLOCK SAVEPOINTIMPFACTORY EXTENDS FactoryBase
VAR
	PRVINSTCOUNT : CAA.COUNT;
	PRVINSTPOOLEXTENDSFACTOR : USINT;
	PRVINSTSIZE : CAA.SIZE;
END_VAR
END_FUNCTION_BLOCK

METHOD CREATE : POINTER TO SavepointImp
VAR_INPUT
	ITFDATA : FBF.IData;
END_VAR
VAR_OUTPUT
	EERROR : FBF.ERROR;
END_VAR
END_METHOD

(* ---- STORAGE.fb ---- *)
FUNCTION_BLOCK STORAGE
VAR
	_HHANDLE : CAA.HANDLE;
	STORAGEENCODING : STO.ENCODING;
	STORAGEISREADONLY : BOOL;
	STORAGELOCKINGSTATE : STO.LOCKING_STATE;
	STORAGENUMOFTABLES : CAA.COUNT;
	STORAGESCHEMAVERSION : DINT;
	STORAGEUSERVERSION : DINT;
	STORAGEVERSION : DINT;
END_VAR
END_FUNCTION_BLOCK

METHOD STORAGECLEAR : STO.ERROR
END_METHOD

METHOD STORAGECLOSE : STO.ERROR
END_METHOD

METHOD STORAGEGETMETRICS : STO.ERROR
VAR_IN_OUT
	MMETRICS : STO.METRICS;
END_VAR
END_METHOD

METHOD STORAGEGETPATH : STO.ERROR
VAR_IN_OUT
	SPATH : CAA.FILENAME;
END_VAR
END_METHOD

METHOD STORAGEOPENFILE : STO.ERROR
VAR_INPUT
	XREADONLY : BOOL := FALSE;
END_VAR
VAR_IN_OUT
	SPATH : CAA.FILENAME;
END_VAR
END_METHOD

METHOD STORAGEREORG : STO.ERROR
END_METHOD

METHOD TABLEOPEN : STO.ITable
VAR_INPUT
	IDTABLE : CAA.IDENT;
END_VAR
VAR_OUTPUT
	EERROR : STO.ERROR;
END_VAR
END_METHOD

METHOD TRANSACTIONBEGIN : STO.ITransaction
VAR_INPUT
	EMODE : STO.TRANSACTION_MODE;
END_VAR
VAR_OUTPUT
	EERROR : STO.ERROR;
END_VAR
END_METHOD

METHOD UTILITYGETCURRENTDATEANDTIME : STO.INT64
VAR_OUTPUT
	EERROR : STO.ERROR;
END_VAR
END_METHOD

METHOD UTILITYRANDOMNESS : STO.ERROR
VAR_INPUT
	SZSIZE : CAA.SIZE;
	PDATA : CAA.PVOID;
END_VAR
END_METHOD

METHOD STORAGEEXECUTESTATEMENT : STO.ERROR
VAR_IN_OUT
	SSTATEMENT : STO.SQLSTATEMENT;
END_VAR
END_METHOD

METHOD STORAGEGETINDEXID : STO.ERROR
VAR_OUTPUT
	IDINDEX : CAA.IDENT;
END_VAR
VAR_IN_OUT
	SINDEX : STRING;
	STABLE : STRING;
END_VAR
END_METHOD

METHOD STORAGEGETTABLEID : STO.ERROR
VAR_OUTPUT
	IDTABLE : CAA.IDENT;
END_VAR
VAR_IN_OUT
	STABLE : STRING;
END_VAR
END_METHOD

(* ---- STORAGEFACTORY.fb ---- *)
FUNCTION_BLOCK STORAGEFACTORY
VAR
	_FACCURSOR : CursorImpFactory;
	_FACROW : RowImpFactory;
	_FACROWPLANCHET : RowPlanchetImpFactory;
	_FACSAVEPOINT : SavepointImpFactory;
	_FACTABLE : TableImpFactory;
	_FACTRANSACTION : TransactionImpFactory;
END_VAR
END_FUNCTION_BLOCK

METHOD CREATECURSOR : STO.ICursor
VAR_INPUT
	HCURSOR : CAA.HANDLE;
	ITFTABLE : STO.ITable;
END_VAR
VAR_OUTPUT
	EERROR : STO.ERROR;
END_VAR
END_METHOD

METHOD CREATEROW : STO.IRow
VAR_INPUT
	HROW : CAA.HANDLE;
	ITFTABLE : STO.ITable;
END_VAR
VAR_OUTPUT
	EERROR : STO.ERROR;
END_VAR
END_METHOD

METHOD CREATEROWPLANCHET : STO.IRowPlanchet
VAR_INPUT
	HROWPLANCHET : CAA.HANDLE;
	ITFTABLE : STO.ITable;
END_VAR
VAR_OUTPUT
	EERROR : STO.ERROR;
END_VAR
END_METHOD

METHOD CREATESAVEPOINT : STO.ISavepoint
VAR_INPUT
	HSAVEPOINT : CAA.HANDLE;
	ITFTRANSACTION : STO.ITransaction;
END_VAR
VAR_OUTPUT
	EERROR : STO.ERROR;
END_VAR
END_METHOD

METHOD CREATETABLE : STO.ITable
VAR_INPUT
	HTABLE : CAA.HANDLE;
	ITFSTORAGE : STO.IStorage;
END_VAR
VAR_OUTPUT
	EERROR : STO.ERROR;
END_VAR
END_METHOD

METHOD CREATETRANSACTION : STO.ITransaction
VAR_INPUT
	HTRANSACTION : TRANSACTION;
	ITFSTORAGE : STO.IStorage;
END_VAR
VAR_OUTPUT
	EERROR : STO.ERROR;
END_VAR
END_METHOD

(* ---- TABLEIMP.fb ---- *)
FUNCTION_BLOCK TABLEIMP EXTENDS InstanceBase
VAR
	_HHANDLE : CAA.HANDLE;
	_ITFSTORAGE : STO.IStorage;
	_EERROR : STO.ERROR;
	LASTERROR : STO.ERROR;
	TABLEID : CAA.IDENT;
	TABLENUMOFCOLUMNS : CAA.COUNT;
	TABLENUMOFINDEXES : CAA.COUNT;
	TABLENUMOFROWS : CAA.COUNT;
	TABLESTORAGE : STO.IStorage;
END_VAR
END_FUNCTION_BLOCK

METHOD ROWDUPLICATE : STO.IRowPlanchet
VAR_INPUT
	IDROW : CAA.IDENT;
END_VAR
VAR_OUTPUT
	EERROR : STO.ERROR;
END_VAR
END_METHOD

METHOD ROWSELECT : STO.IRow
VAR_INPUT
	IDROW : CAA.IDENT;
END_VAR
VAR_OUTPUT
	EERROR : STO.ERROR;
END_VAR
END_METHOD

METHOD PRVINSTINIT : FBF.ERROR
VAR_INPUT
	ITFDATA : FBF.IData;
END_VAR
END_METHOD

METHOD ROWDELETE2 : STO.ERROR
VAR_INPUT
	IDROW : LINT;
END_VAR
END_METHOD

METHOD TABLECLOSE : STO.ERROR
END_METHOD

METHOD GETMINMAXROWIDS : STO.ERROR
VAR_OUTPUT
	IDROWMIN : LINT;
	IDROWMAX : LINT;
END_VAR
END_METHOD

METHOD ROWDELETE : STO.ERROR
VAR_INPUT
	IDROW : CAA.IDENT;
END_VAR
END_METHOD

METHOD ROWCREATE : STO.IRowPlanchet
VAR_OUTPUT
	EERROR : STO.ERROR;
END_VAR
END_METHOD

METHOD TABLECLEAR : STO.ERROR
END_METHOD

METHOD CURSOROPEN : STO.ICursor
VAR_INPUT
	IDINDEX : CAA.IDENT;
	XREADONLY : BOOL;
END_VAR
VAR_OUTPUT
	EERROR : STO.ERROR;
END_VAR
END_METHOD

(* ---- TABLEIMPFACTORY.fb ---- *)
FUNCTION_BLOCK TABLEIMPFACTORY EXTENDS FactoryBase
VAR
	PRVINSTCOUNT : CAA.COUNT;
	PRVINSTPOOLEXTENDSFACTOR : USINT;
	PRVINSTSIZE : CAA.SIZE;
END_VAR
END_FUNCTION_BLOCK

METHOD CREATE : POINTER TO TableImp
VAR_INPUT
	ITFDATA : FBF.IData;
END_VAR
VAR_OUTPUT
	EERROR : FBF.ERROR;
END_VAR
END_METHOD

(* ---- TRANSACTIONIMP.fb ---- *)
FUNCTION_BLOCK TRANSACTIONIMP EXTENDS InstanceBase
VAR
	_HHANDLE : CAA.HANDLE;
	_ITFSTORAGE : STO.IStorage;
	TRANSACTIONSTORAGE : STO.IStorage;
END_VAR
END_FUNCTION_BLOCK

METHOD TRANSACTIONCOMMIT : STO.ERROR
END_METHOD

METHOD TRANSACTIONROLLBACK : STO.ERROR
END_METHOD

METHOD TRANSACTIONSETSAVEPOINT : STO.ISavepoint
VAR_OUTPUT
	EERROR : STO.ERROR;
END_VAR
END_METHOD

METHOD PRVINSTINIT : FBF.ERROR
VAR_INPUT
	ITFDATA : FBF.IData;
END_VAR
END_METHOD

(* ---- TRANSACTIONIMPFACTORY.fb ---- *)
FUNCTION_BLOCK TRANSACTIONIMPFACTORY EXTENDS FactoryBase
VAR
	PRVINSTCOUNT : CAA.COUNT;
	PRVINSTPOOLEXTENDSFACTOR : USINT;
	PRVINSTSIZE : CAA.SIZE;
END_VAR
END_FUNCTION_BLOCK

METHOD CREATE : POINTER TO TransactionImp
VAR_INPUT
	ITFDATA : FBF.IData;
END_VAR
VAR_OUTPUT
	EERROR : FBF.ERROR;
END_VAR
END_METHOD
